Staubli VAL3: initDataBase.pgx

program initDataBase()
begin
  db:nStep0=10
  db:nStep1=10
  db:nStep2=10
  db:nStep3=10
  //
  db:tFlange.trsf={0,0,0,0,0,0}
  db:trOffset={0,0,10,0,0,0}
  //
  db:mSpeed_C_blend.tvel=250
  db:mSpeed_C_blend.blend=Cartesian
  db:mSpeed_C_blend.leave=0
  db:mSpeed_C_blend.reach=0
  //
  db:mSpeed_J_blend.tvel=250
  db:mSpeed_J_blend.blend=joint
  db:mSpeed_J_blend.leave=5
  db:mSpeed_J_blend.reach=5
  //
  db:mSlow.tvel=30
  db:mSlow.blend=Cartesian
  db:mSlow.leave=0
  db:mSlow.reach=0
  //
  db:cConfigSame={ssame,esame,wsame}
  //
  //pTeach1.trsf={0,0,0,0,0,0}
  db:pTeach1.config={ssame,esame,wsame}
  //pTeach2.trsf={0,0,0,0,0,0}
  db:pTeach2.config={ssame,esame,wsame}
  //pTeach3.trsf={0,0,0,0,0,0}
  db:pTeach3.config={ssame,esame,wsame}
  //pTeach4.trsf={0,0,0,0,0,0}
  db:pTeach4.config={ssame,esame,wsame}
  //pTeach5.trsf={0,0,0,0,0,0}
  db:pTeach5.config={ssame,esame,wsame}
  //pTeach6.trsf={0,0,0,0,0,0}
  db:pTeach6.config={ssame,esame,wsame}
  //pTeach6.trsf={0,0,0,0,0,0}
  db:pTeach7.config={ssame,esame,wsame}
  //
  //pAdjustXY_2_1.trsf={0,0,0,0,0,0}
  db:pAdjustXY_2_1.config={ssame,esame,wsame}
  //pAdjustXY_2_2.trsf={0,0,0,0,0,0}
  db:pAdjustXY_2_2.config={ssame,esame,wsame}
  //pAdjustXY_3_1.trsf={0,0,0,0,0,0}
  db:pAdjustXY_3_1.config={ssame,esame,wsame}
  //pAdjustXY_3_2.trsf={0,0,0,0,0,0}
  db:pAdjustXY_3_2.config={ssame,esame,wsame}
  //pAdjustXY_3_3.trsf={0,0,0,0,0,0}
  db:pAdjustXY_3_3.config={ssame,esame,wsame}
  //pAdjustZ_2_1.trsf={0,0,0,0,0,0}
  db:pAdjustZ_2_1.config={ssame,esame,wsame}
  //pAdjustZ_2_2.trsf={0,0,0,0,0,0}
  db:pAdjustZ_2_2.config={ssame,esame,wsame}
  //
  db:bTeach1=false
  db:bTeach2=false
  db:bTeach3=false
  db:bTeach4=false
  db:bTeach5=false
  db:bTeach6=false
  db:bTeach7=false
  //
  db:bAdjustXY_2_1=false
  db:bAdjustXY_2_2=false
  db:bAdjustXY_3_1=false
  db:bAdjustXY_3_2=false
  db:bAdjustXY_3_3=false
  db:bAdjustZ_2_1=false
  db:bAdjustZ_2_2=false
  //
  db:sLanguageM=""
  db:sCbxLanguage=""
  db:sCbxMounting=""
end
